INTERFACE I_LevelSensor EXTENDS __SYSTEM.IQueryInterface

PROPERTY Level : REAL
GET
END_GET
END_PROPERTY

PROPERTY IsValid : BOOL
GET
END_GET
END_PROPERTY

END_INTERFACE

(* stored: Version 1.1.0.1
   Itf I_LevelSensor: Id {d0b6623f-94bb-4398-810a-73c95ba7647d}
   Property Level: Id {6bcab137-6eb8-43d8-a561-ab7034a300b0}
   Get Get: Id {4b37a827-031a-4b10-a052-e46b9ebea635}
   Property IsValid: Id {6a949da8-fdef-41a0-8d20-8cae3d78d7dc}
   Get Get: Id {ece6091c-8d84-4c88-87f2-f806a8759538} *)
